// TIA Portal V21 export
FUNCTION_BLOCK "FB_AnaShared"   // FB16, SCL
TITLE = Analyzer: instance shared by two OBs
{ S7_Optimized_Access := 'TRUE' }
// Rule C26l: the instance IDB_AnaShared is called from OB_Main and from OB_Cyclic100ms
// stored: MemoryReserve 100, SetENOAutomatically false
   VAR_INPUT
      Pulse : Bool;   // Count pulse
   END_VAR
   VAR_OUTPUT
      Count : Int;   // Number of pulses
   END_VAR
   VAR
      PulseEdge { S7_SetPoint := 'True'} : R_TRIG;   // Edge of the pulse
   END_VAR
BEGIN

       #PulseEdge(CLK := #Pulse);
       IF #PulseEdge.Q THEN
           #Count := #Count + 1;
       END_IF;
END_FUNCTION_BLOCK
